Staubli VAL3: start.pgx

public program start()
begin
  if prog:libLoad("./TgtProg")!=0
    logMsg("Error Loading RoboDK library")
    popUpMsg("Error Loading RoboDK library")
  endIf
  wait(taskStatus("loading")==-1)
  taskCreate "loading",10,loadNextOne("./TgtProg2")
  call prog:start()

  if prog:libLoad("./TgtProg2")!=0
    logMsg("Error Loading RoboDK library")
    popUpMsg("Error Loading RoboDK library")
  endIf
  wait(taskStatus("loading")==-1)
  call prog:start()


end
